TYPE ST_EL9576 :
STRUCT
    sTerminalName : STRING(200) := 'EL9576 | Brake Chopper Terminal';

    stTerminalInfo : ST_Terminal_Info;
END_STRUCT
END_TYPE

(* stored: Version 1.1.0.1, ProductVersion 3.1.4026.18
   DUT ST_EL9576: Id {2aa121e2-110b-404c-8b02-49035f0fac4e} *)
